(* IEC 61131-3 sources: llm-plc-st-eval/data/processed_v2_primera/gpt-4o/I1/few_shot, 3 files *)

(* ---- ejec_1.st ---- *)
FUNCTION_BLOCK FB_Semaforo
VAR_INPUT
    habilitado : BOOL; (* Habilita el funcionamiento del semáforo *)
END_VAR
VAR_OUTPUT
    luzV : BOOL; (* Luz verde del semáforo *)
    luzA : BOOL; (* Luz amarilla del semáforo *)
    luzR : BOOL; (* Luz roja del semáforo *)
END_VAR
VAR
    tCiclo : TON; (* Temporizador para el ciclo del semáforo *)
    tIntermitente : TON; (* Temporizador para el amarillo intermitente *)
    estado : INT; (* Estado actual del semáforo *)
END_VAR

(* Inicialización de variables *)
IF NOT habilitado THEN
    (* Modo amarillo intermitente *)
    tIntermitente(IN := TRUE, PT := T#1S);
    luzV := FALSE;
    luzR := FALSE;
    luzA := tIntermitente.Q;
    estado := 0; (* Reinicia el estado para cuando se habilite de nuevo *)
ELSE
    (* Modo ciclo normal del semáforo *)
    tIntermitente(IN := FALSE);
    CASE estado OF
        0: (* Luz verde *)
            tCiclo(IN := TRUE, PT := T#20S);
            luzV := TRUE;
            luzA := FALSE;
            luzR := FALSE;
            IF tCiclo.Q THEN
                estado := 1;
                tCiclo(IN := FALSE);
            END_IF;
        1: (* Luz amarilla *)
            tCiclo(IN := TRUE, PT := T#4S);
            luzV := FALSE;
            luzA := TRUE;
            luzR := FALSE;
            IF tCiclo.Q THEN
                estado := 2;
                tCiclo(IN := FALSE);
            END_IF;
        2: (* Luz roja *)
            tCiclo(IN := TRUE, PT := T#15S);
            luzV := FALSE;
            luzA := FALSE;
            luzR := TRUE;
            IF tCiclo.Q THEN
                estado := 0;
                tCiclo(IN := FALSE);
            END_IF;
    END_CASE;
END_IF;
END_FUNCTION_BLOCK

(* ---- ejec_2.st ---- *)
FUNCTION_BLOCK FB_Semaforo
VAR_INPUT
    habilitado : BOOL; (* Habilitacion del semaforo *)
END_VAR
VAR_OUTPUT
    luzV : BOOL; (* Luz verde *)
    luzA : BOOL; (* Luz amarilla *)
    luzR : BOOL; (* Luz roja *)
END_VAR
VAR
    tCiclo : TON; (* Temporizador para el ciclo del semaforo *)
    tIntermitente : TON; (* Temporizador para el amarillo intermitente *)
    estado : INT; (* Estado del semaforo *)
END_VAR

(* Inicializacion de variables *)
IF NOT habilitado THEN
    (* Modo amarillo intermitente *)
    tIntermitente(IN := TRUE, PT := T#1S);
    luzV := FALSE;
    luzR := FALSE;
    luzA := tIntermitente.Q;
    tCiclo(IN := FALSE);
    estado := 0; (* Reiniciar estado al habilitarse de nuevo *)
ELSE
    (* Modo ciclo normal *)
    tIntermitente(IN := FALSE);
    CASE estado OF
        0: (* Luz verde *)
            luzV := TRUE;
            luzA := FALSE;
            luzR := FALSE;
            tCiclo(IN := TRUE, PT := T#20S);
            IF tCiclo.Q THEN
                estado := 1;
                tCiclo(IN := FALSE);
            END_IF
        1: (* Luz amarilla *)
            luzV := FALSE;
            luzA := TRUE;
            luzR := FALSE;
            tCiclo(IN := TRUE, PT := T#4S);
            IF tCiclo.Q THEN
                estado := 2;
                tCiclo(IN := FALSE);
            END_IF
        2: (* Luz roja *)
            luzV := FALSE;
            luzA := FALSE;
            luzR := TRUE;
            tCiclo(IN := TRUE, PT := T#15S);
            IF tCiclo.Q THEN
                estado := 0;
                tCiclo(IN := FALSE);
            END_IF
    END_CASE
END_IF
END_FUNCTION_BLOCK

(* ---- ejec_3.st ---- *)
FUNCTION_BLOCK FB_Semaforo
VAR_INPUT
    habilitado : BOOL; (* Habilitacion del semaforo *)
END_VAR
VAR_OUTPUT
    luzV : BOOL; (* Luz verde *)
    luzA : BOOL; (* Luz amarilla *)
    luzR : BOOL; (* Luz roja *)
END_VAR
VAR
    tVerde : TON; (* Temporizador para luz verde *)
    tAmarillo : TON; (* Temporizador para luz amarilla *)
    tRojo : TON; (* Temporizador para luz roja *)
    tIntermitente : TON; (* Temporizador para amarillo intermitente *)
    estado : INT; (* Estado del semaforo *)
END_VAR

(* Logica del semaforo *)
IF habilitado THEN
    CASE estado OF
        0: (* Estado verde *)
            tVerde(IN := TRUE, PT := T#20S);
            luzV := tVerde.Q;
            luzA := FALSE;
            luzR := FALSE;
            IF tVerde.Q THEN
                tVerde(IN := FALSE);
                estado := 1;
            END_IF;
        1: (* Estado amarillo *)
            tAmarillo(IN := TRUE, PT := T#4S);
            luzV := FALSE;
            luzA := tAmarillo.Q;
            luzR := FALSE;
            IF tAmarillo.Q THEN
                tAmarillo(IN := FALSE);
                estado := 2;
            END_IF;
        2: (* Estado rojo *)
            tRojo(IN := TRUE, PT := T#15S);
            luzV := FALSE;
            luzA := FALSE;
            luzR := tRojo.Q;
            IF tRojo.Q THEN
                tRojo(IN := FALSE);
                estado := 0;
            END_IF;
    END_CASE;
ELSE
    (* Estado amarillo intermitente *)
    tIntermitente(IN := TRUE, PT := T#1S);
    luzV := FALSE;
    luzA := tIntermitente.Q;
    luzR := FALSE;
    IF tIntermitente.Q THEN
        tIntermitente(IN := FALSE);
    END_IF;
    estado := 0; (* Reinicia el ciclo al habilitarse *)
END_IF;
END_FUNCTION_BLOCK
